// TIA Portal V20 export
Screen "Pop-up_ControlOnOff_Popup"  310x143
  ScreenItem "Background" at 0,0 size 310x143  Type=HmiRectangle
  ScreenItem "Overview_SafetyDialog" at 1,1 size 308x25  Type=HmiTextBox
  ScreenItem "Descr_ONOFF" at 3,26 size 184x25  Type=HmiTextBox
  ScreenItem "Button_Power_Off" at 110,73 size 90x60  Type=HmiButton
  ScreenItem "Button_Close" at 219,1 size 90x59  Type=HmiButton
  ScreenItem "Button_Cancel" at 210,73 size 90x60  Type=HmiButton
  ScreenItem "Button_Power_On" at 10,73 size 90x60  Type=HmiButton
